ABB RAPID module: SplitTest_1.mod

%%%
  VERSION:1
  LANGUAGE:ENGLISH
%%%
MODULE MOD_Tmp2

	PROC Prg_Tmp2()

		MoveL [[315.779,-74.668,245.881],[0.09884449,0.01379658,0.99324025,0.05927254],[-1,0,-1,0],[9E+09,9E+09,9E+09,9E+09,9E+09,9E+09]],v200,z1,Tool1 \WObj:=Frame2;
		MoveL [[284.148,-86.783,243.844],[0.09359571,0.04936652,0.99254150,0.06053239],[-1,0,-1,0],[9E+09,9E+09,9E+09,9E+09,9E+09,9E+09]],v200,z1,Tool1 \WObj:=Frame2;
		MoveL [[315.779,-74.668,245.881],[0.09884449,0.01379658,0.99324025,0.05927254],[-1,0,-1,0],[9E+09,9E+09,9E+09,9E+09,9E+09,9E+09]],v200,z1,Tool1 \WObj:=Frame2;
		MoveL [[284.148,-86.783,243.844],[0.09359571,0.04936652,0.99254150,0.06053239],[-1,0,-1,0],[9E+09,9E+09,9E+09,9E+09,9E+09,9E+09]],v200,z1,Tool1 \WObj:=Frame2;
		MoveL [[315.779,-74.668,245.881],[0.09884449,0.01379658,0.99324025,0.05927254],[-1,0,-1,0],[9E+09,9E+09,9E+09,9E+09,9E+09,9E+09]],v200,z1,Tool1 \WObj:=Frame2;
		MoveL [[284.148,-86.783,243.844],[0.09359571,0.04936652,0.99254150,0.06053239],[-1,0,-1,0],[9E+09,9E+09,9E+09,9E+09,9E+09,9E+09]],v200,z1,Tool1 \WObj:=Frame2;
		MoveL [[315.779,-74.668,245.881],[0.09884449,0.01379658,0.99324025,0.05927254],[-1,0,-1,0],[9E+09,9E+09,9E+09,9E+09,9E+09,9E+09]],v200,z1,Tool1 \WObj:=Frame2;
		MoveL [[284.148,-86.783,243.844],[0.09359571,0.04936652,0.99254150,0.06053239],[-1,0,-1,0],[9E+09,9E+09,9E+09,9E+09,9E+09,9E+09]],v200,z1,Tool1 \WObj:=Frame2;
		MoveL [[315.779,-74.668,245.881],[0.09884449,0.01379658,0.99324025,0.05927254],[-1,0,-1,0],[9E+09,9E+09,9E+09,9E+09,9E+09,9E+09]],v200,z1,Tool1 \WObj:=Frame2;
		MoveL [[284.148,-86.783,243.844],[0.09359571,0.04936652,0.99254150,0.06053239],[-1,0,-1,0],[9E+09,9E+09,9E+09,9E+09,9E+09,9E+09]],v200,z1,Tool1 \WObj:=Frame2;
		MoveL [[315.779,-74.668,245.881],[0.09884449,0.01379658,0.99324025,0.05927254],[-1,0,-1,0],[9E+09,9E+09,9E+09,9E+09,9E+09,9E+09]],v200,z1,Tool1 \WObj:=Frame2;
		MoveL [[284.148,-86.783,243.844],[0.09359571,0.04936652,0.99254150,0.06053239],[-1,0,-1,0],[9E+09,9E+09,9E+09,9E+09,9E+09,9E+09]],v200,z1,Tool1 \WObj:=Frame2;
		MoveL [[315.779,-74.668,245.881],[0.09884449,0.01379658,0.99324025,0.05927254],[-1,0,-1,0],[9E+09,9E+09,9E+09,9E+09,9E+09,9E+09]],v200,z1,Tool1 \WObj:=Frame2;
		MoveL [[284.148,-86.783,243.844],[0.09359571,0.04936652,0.99254150,0.06053239],[-1,0,-1,0],[9E+09,9E+09,9E+09,9E+09,9E+09,9E+09]],v200,z1,Tool1 \WObj:=Frame2;
		MoveL [[315.779,-74.668,245.881],[0.09884449,0.01379658,0.99324025,0.05927254],[-1,0,-1,0],[9E+09,9E+09,9E+09,9E+09,9E+09,9E+09]],v200,z1,Tool1 \WObj:=Frame2;

	ENDPROC

ENDMODULE
